(* Logix 5000 project; controller TFF vendor 1 type 14 code 107 rev 34.11; software revision 34.03; part 31 of 36 *)
(* tags used below, declared in another part *)
   FlowPath : FlowPath[64];   // Flow Path Array
   FlowPathControl : FlowPathControl;   // Flow Path Control
   Options : Options;   // Options List
   PCV001_Control : PCV_Control;   // PCV001 Control UDT
   PipeAnimation : PipeAnimation;   // HMI Pipe Animation Array
   XV001 : ALIAS FOR Valve[0];   // XV001
   XV002 : ALIAS FOR Valve[1];   // XV002
   XV003 : ALIAS FOR Valve[2];   // XV003
   XV004 : ALIAS FOR Valve[3];   // XV004
   XV005 : ALIAS FOR Valve[4];   // XV005
   XV006 : ALIAS FOR Valve[19];
   XV007 : ALIAS FOR Valve[20];
   XV401 : ALIAS FOR Valve[6];   // XV401
   XV402 : ALIAS FOR Valve[7];   // XV402
   XV403 : ALIAS FOR Valve[15];
   XV404 : ALIAS FOR Valve[16];
   XV405 : ALIAS FOR Valve[17];
   XV406 : ALIAS FOR Valve[18];
   XV411 : ALIAS FOR Valve[8];   // XV411
   XV421 : ALIAS FOR Valve[9];   // XV421
   XV431 : ALIAS FOR Valve[10];   // XV431
   XV441 : ALIAS FOR Valve[11];   // XV441
   XV901 : ALIAS FOR Valve[14];   // XV901
(* Process, continued *)

ROUTINE PipeAnimationControl   (* ladder *)
// Pipework Animation Routine
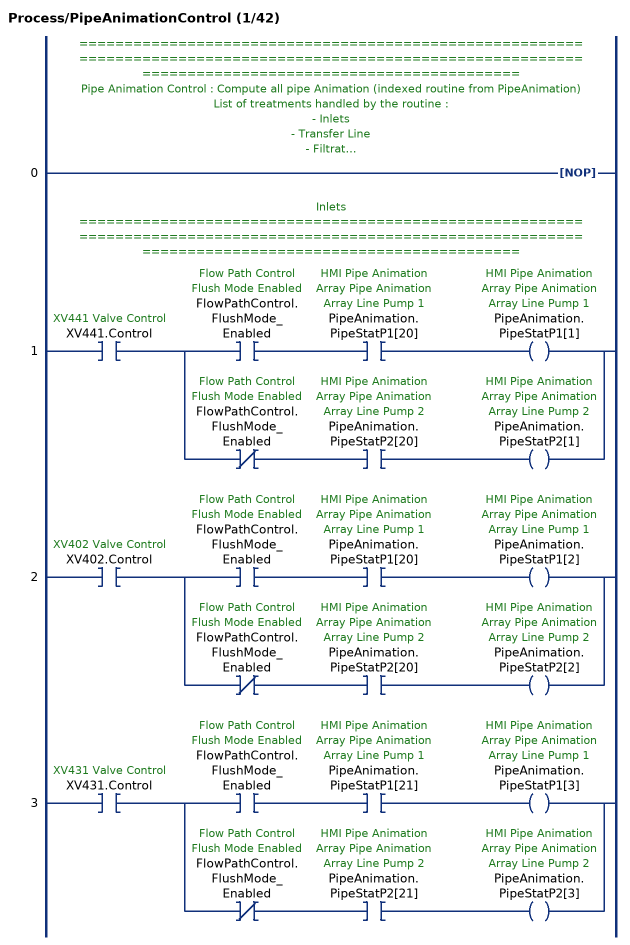
   // ==========================================================================================================================================================
   //                                                                                        Pipe Animation Control : Compute all pipe Animation (indexed routine from PipeAnimation)
   //                                                     List of treatments handled by the routine :
   //                                                          - Inlets
   //                                                          - Transfer Line
   //                                                          - Filtrate
   //                                                          - Flush
   //                                                     -----------------------------------------------------------------------------------------------------------------------------------------------------
   //                                                     History
   //                                                          2019-AUG-13 - Actemium - B. Roch - Initial version for Candidate Release 3.00.00.00.a
   //                                                          2020-OCT-01 - Merck - Q. Spindler - Modifications for Candidate Release 3.00.00.01.a
   //                                                   - Change pipe animation to add Closed Flowpath option
   // - Lock Frontal filtration flowpath
   // ========================================================================================================================================================
   0: NOP();
   // Inlets
   // ==========================================================================================================================================================
   1: XIC(XV441.Control)[XIC(FlowPathControl.FlushMode_Enabled) XIC(PipeAnimation.PipeStatP1[20]) OTE(PipeAnimation.PipeStatP1[1]) ,XIO(FlowPathControl.FlushMode_Enabled) XIC(PipeAnimation.PipeStatP2[20]) OTE(PipeAnimation.PipeStatP2[1]) ];
   2: XIC(XV402.Control)[XIC(FlowPathControl.FlushMode_Enabled) XIC(PipeAnimation.PipeStatP1[20]) OTE(PipeAnimation.PipeStatP1[2]) ,XIO(FlowPathControl.FlushMode_Enabled) XIC(PipeAnimation.PipeStatP2[20]) OTE(PipeAnimation.PipeStatP2[2]) ];
   3: XIC(XV431.Control)[XIC(FlowPathControl.FlushMode_Enabled) XIC(PipeAnimation.PipeStatP1[21]) OTE(PipeAnimation.PipeStatP1[3]) ,XIO(FlowPathControl.FlushMode_Enabled) XIC(PipeAnimation.PipeStatP2[21]) OTE(PipeAnimation.PipeStatP2[3]) ];
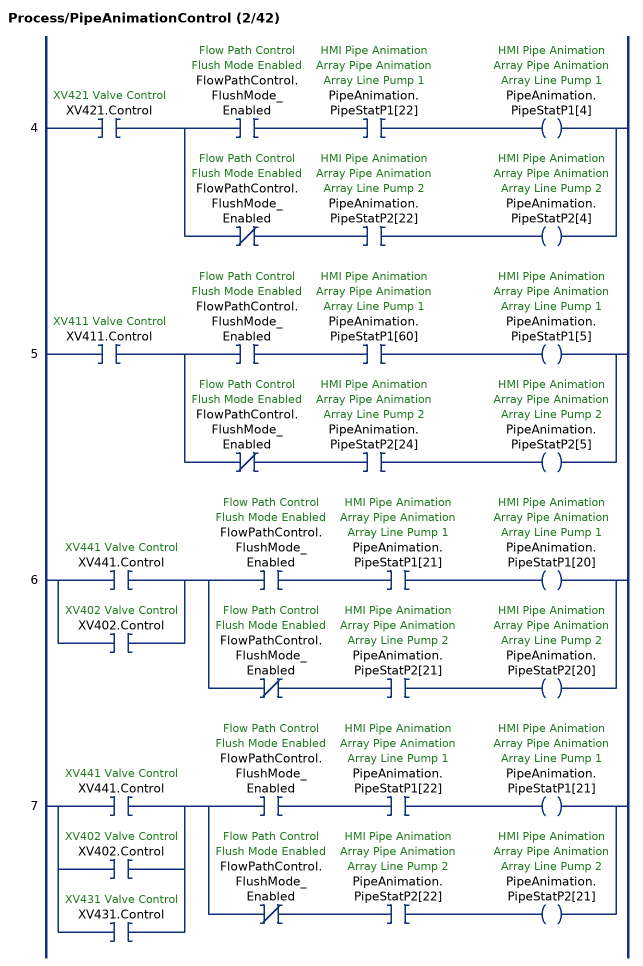
   4: XIC(XV421.Control)[XIC(FlowPathControl.FlushMode_Enabled) XIC(PipeAnimation.PipeStatP1[22]) OTE(PipeAnimation.PipeStatP1[4]) ,XIO(FlowPathControl.FlushMode_Enabled) XIC(PipeAnimation.PipeStatP2[22]) OTE(PipeAnimation.PipeStatP2[4]) ];
   5: XIC(XV411.Control)[XIC(FlowPathControl.FlushMode_Enabled) XIC(PipeAnimation.PipeStatP1[60]) OTE(PipeAnimation.PipeStatP1[5]) ,XIO(FlowPathControl.FlushMode_Enabled) XIC(PipeAnimation.PipeStatP2[24]) OTE(PipeAnimation.PipeStatP2[5]) ];
   6: [XIC(XV441.Control) ,XIC(XV402.Control) ][XIC(FlowPathControl.FlushMode_Enabled) XIC(PipeAnimation.PipeStatP1[21]) OTE(PipeAnimation.PipeStatP1[20]) ,XIO(FlowPathControl.FlushMode_Enabled) XIC(PipeAnimation.PipeStatP2[21]) OTE(PipeAnimation.PipeStatP2[20]) ];
   7: [XIC(XV441.Control) ,XIC(XV402.Control) ,XIC(XV431.Control) ][XIC(FlowPathControl.FlushMode_Enabled) XIC(PipeAnimation.PipeStatP1[22]) OTE(PipeAnimation.PipeStatP1[21]) ,XIO(FlowPathControl.FlushMode_Enabled) XIC(PipeAnimation.PipeStatP2[22]) OTE(PipeAnimation.PipeStatP2[21]) ];
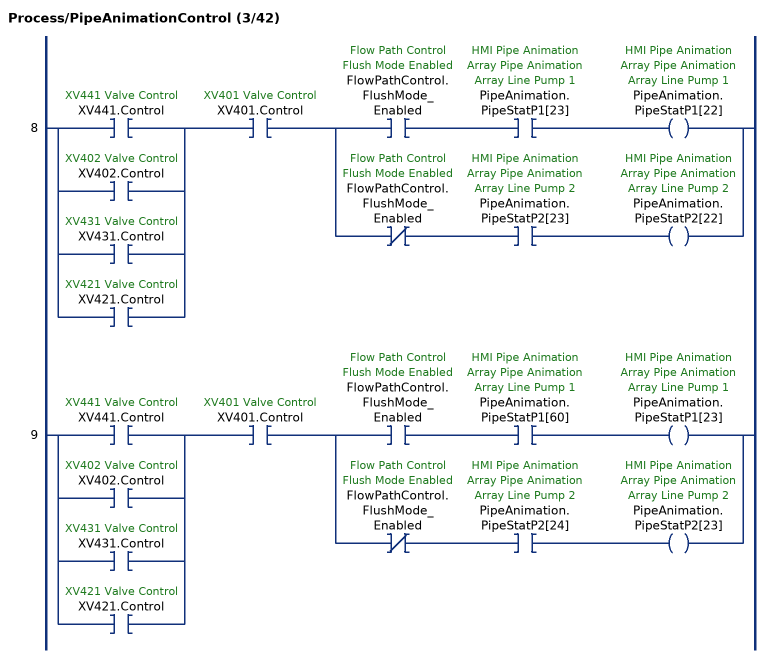
   8: [XIC(XV441.Control) ,XIC(XV402.Control) ,XIC(XV431.Control) ,XIC(XV421.Control) ]XIC(XV401.Control)[XIC(FlowPathControl.FlushMode_Enabled) XIC(PipeAnimation.PipeStatP1[23]) OTE(PipeAnimation.PipeStatP1[22]) ,XIO(FlowPathControl.FlushMode_Enabled) XIC(PipeAnimation.PipeStatP2[23]) OTE(PipeAnimation.PipeStatP2[22]) ];
   9: [XIC(XV441.Control) ,XIC(XV402.Control) ,XIC(XV431.Control) ,XIC(XV421.Control) ]XIC(XV401.Control)[XIC(FlowPathControl.FlushMode_Enabled) XIC(PipeAnimation.PipeStatP1[60]) OTE(PipeAnimation.PipeStatP1[23]) ,XIO(FlowPathControl.FlushMode_Enabled) XIC(PipeAnimation.PipeStatP2[24]) OTE(PipeAnimation.PipeStatP2[23]) ];
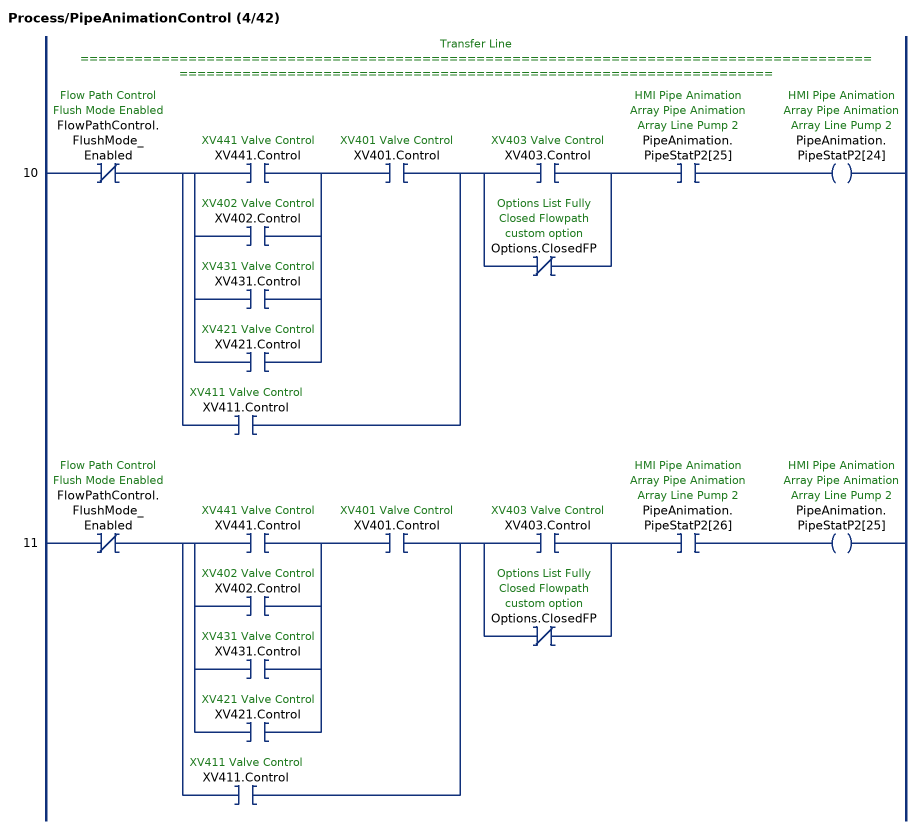
   // Transfer Line
   // ==========================================================================================================================================================
   10: XIO(FlowPathControl.FlushMode_Enabled)[[XIC(XV441.Control) ,XIC(XV402.Control) ,XIC(XV431.Control) ,XIC(XV421.Control) ] XIC(XV401.Control) ,XIC(XV411.Control) ][XIC(XV403.Control) ,XIO(Options.ClosedFP) ]XIC(PipeAnimation.PipeStatP2[25])OTE(PipeAnimation.PipeStatP2[24]);
   11: XIO(FlowPathControl.FlushMode_Enabled)[[XIC(XV441.Control) ,XIC(XV402.Control) ,XIC(XV431.Control) ,XIC(XV421.Control) ] XIC(XV401.Control) ,XIC(XV411.Control) ][XIC(XV403.Control) ,XIO(Options.ClosedFP) ]XIC(PipeAnimation.PipeStatP2[26])OTE(PipeAnimation.PipeStatP2[25]);
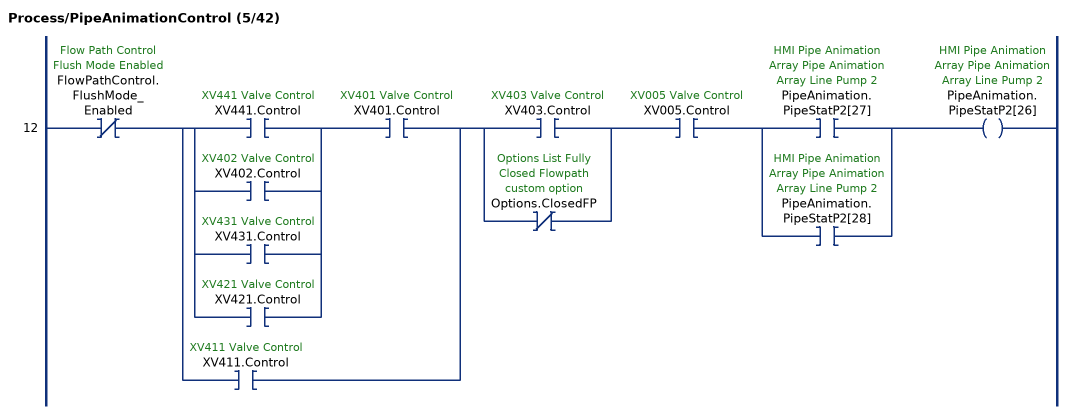
   12: XIO(FlowPathControl.FlushMode_Enabled)[[XIC(XV441.Control) ,XIC(XV402.Control) ,XIC(XV431.Control) ,XIC(XV421.Control) ] XIC(XV401.Control) ,XIC(XV411.Control) ][XIC(XV403.Control) ,XIO(Options.ClosedFP) ]XIC(XV005.Control)[XIC(PipeAnimation.PipeStatP2[27]) ,XIC(PipeAnimation.PipeStatP2[28]) ]OTE(PipeAnimation.PipeStatP2[26]);
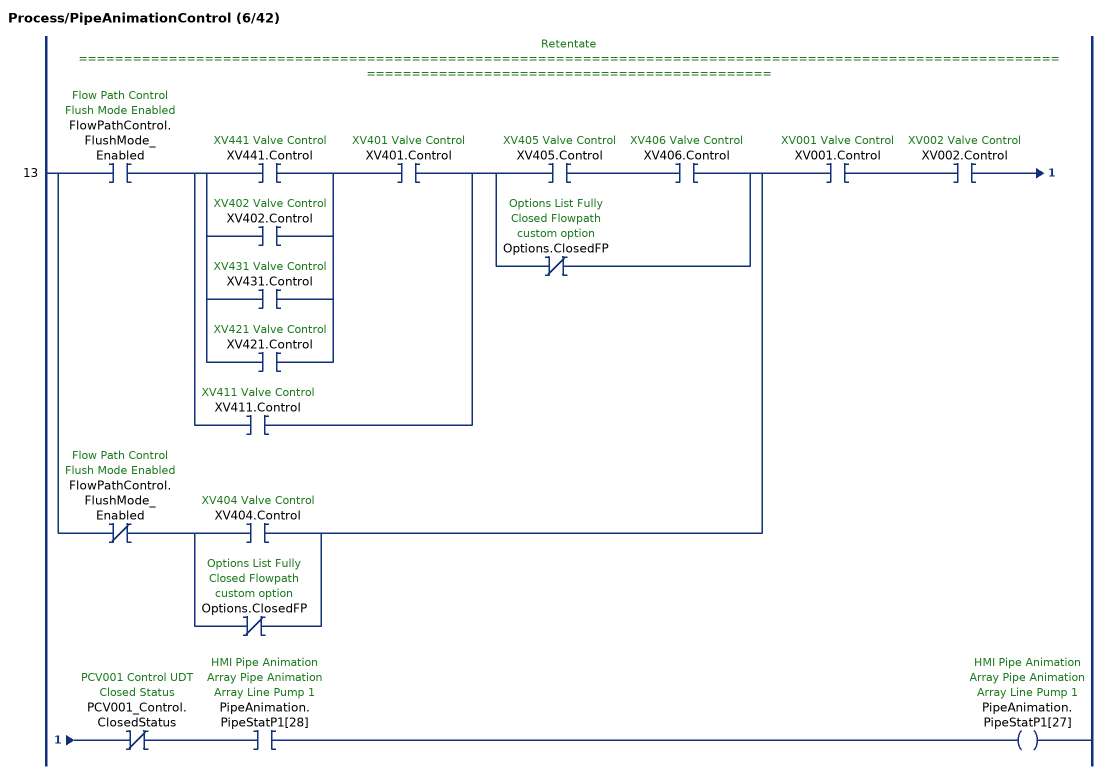
   // Retentate
   // ==========================================================================================================================================================
   13: [XIC(FlowPathControl.FlushMode_Enabled) [[XIC(XV441.Control) ,XIC(XV402.Control) ,XIC(XV431.Control) ,XIC(XV421.Control) ] XIC(XV401.Control) ,XIC(XV411.Control) ] [XIC(XV405.Control) XIC(XV406.Control) ,XIO(Options.ClosedFP) ] ,XIO(FlowPathControl.FlushMode_Enabled) [XIC(XV404.Control) ,XIO(Options.ClosedFP) ] ]XIC(XV001.Control)XIC(XV002.Control)XIO(PCV001_Control.ClosedStatus)XIC(PipeAnimation.PipeStatP1[28])OTE(PipeAnimation.PipeStatP1[27]);
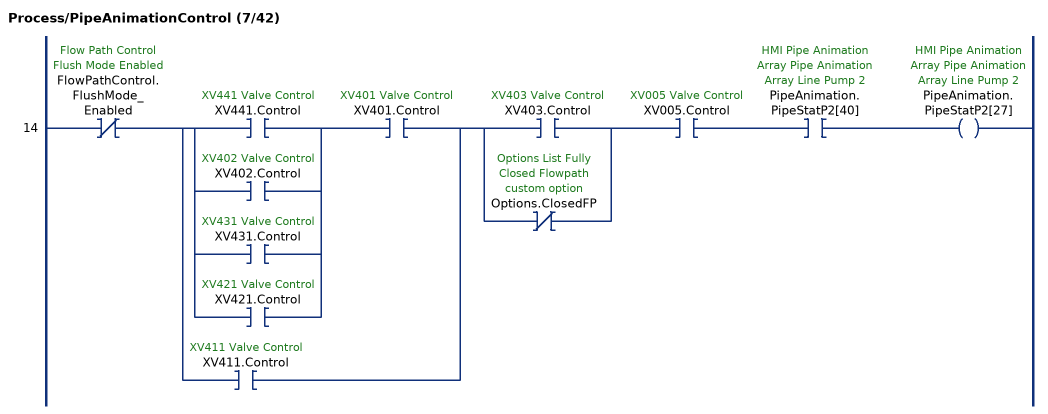
   14: XIO(FlowPathControl.FlushMode_Enabled)[[XIC(XV441.Control) ,XIC(XV402.Control) ,XIC(XV431.Control) ,XIC(XV421.Control) ] XIC(XV401.Control) ,XIC(XV411.Control) ][XIC(XV403.Control) ,XIO(Options.ClosedFP) ]XIC(XV005.Control)XIC(PipeAnimation.PipeStatP2[40])OTE(PipeAnimation.PipeStatP2[27]);
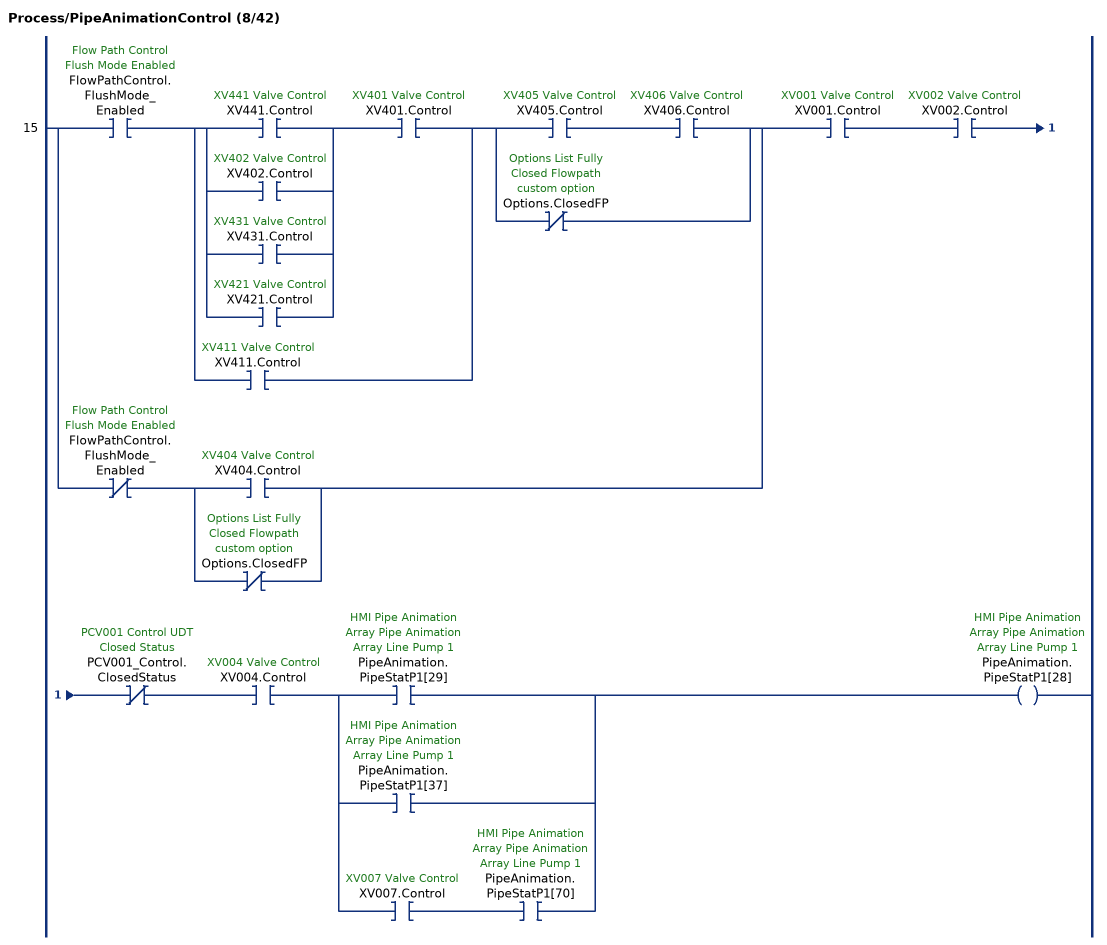
   15: [XIC(FlowPathControl.FlushMode_Enabled) [[XIC(XV441.Control) ,XIC(XV402.Control) ,XIC(XV431.Control) ,XIC(XV421.Control) ] XIC(XV401.Control) ,XIC(XV411.Control) ] [XIC(XV405.Control) XIC(XV406.Control) ,XIO(Options.ClosedFP) ] ,XIO(FlowPathControl.FlushMode_Enabled) [XIC(XV404.Control) ,XIO(Options.ClosedFP) ] ]XIC(XV001.Control)XIC(XV002.Control)XIO(PCV001_Control.ClosedStatus)XIC(XV004.Control)[[XIC(PipeAnimation.PipeStatP1[29]) ,XIC(PipeAnimation.PipeStatP1[37]) ] ,XIC(XV007.Control) XIC(PipeAnimation.PipeStatP1[70]) ]OTE(PipeAnimation.PipeStatP1[28]);
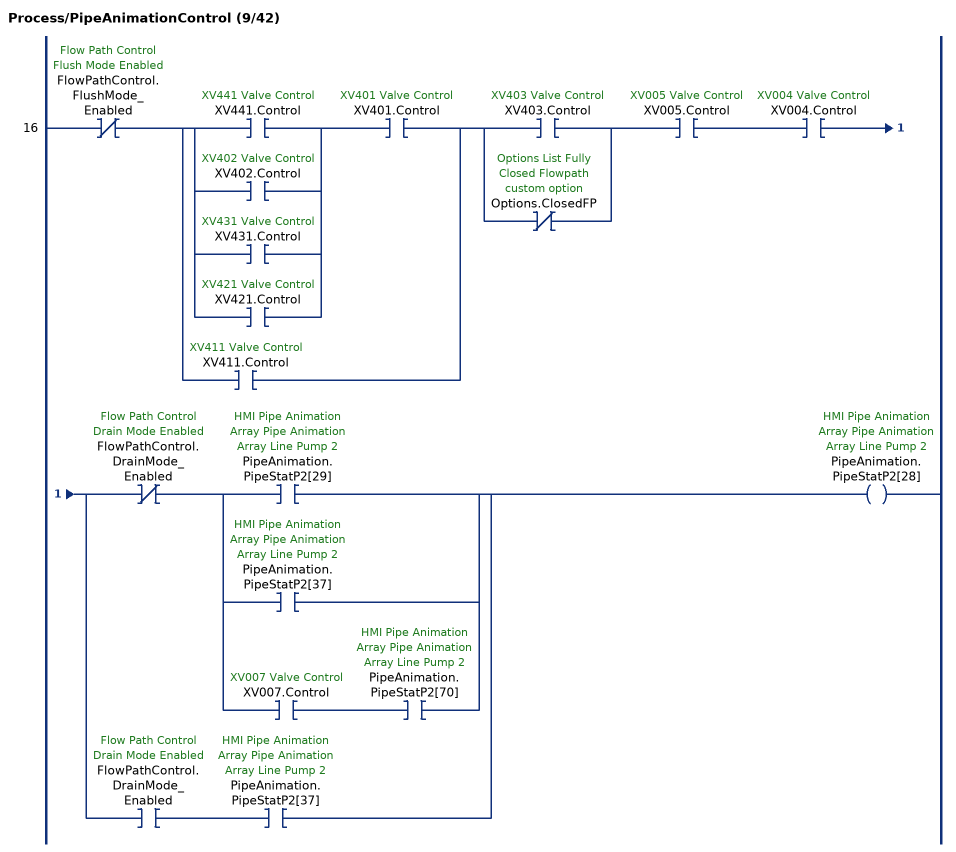
   16: XIO(FlowPathControl.FlushMode_Enabled)[[XIC(XV441.Control) ,XIC(XV402.Control) ,XIC(XV431.Control) ,XIC(XV421.Control) ] XIC(XV401.Control) ,XIC(XV411.Control) ][XIC(XV403.Control) ,XIO(Options.ClosedFP) ]XIC(XV005.Control)XIC(XV004.Control)[XIO(FlowPathControl.DrainMode_Enabled) [[XIC(PipeAnimation.PipeStatP2[29]) ,XIC(PipeAnimation.PipeStatP2[37]) ] ,XIC(XV007.Control) XIC(PipeAnimation.PipeStatP2[70]) ] ,XIC(FlowPathControl.DrainMode_Enabled) XIC(PipeAnimation.PipeStatP2[37]) ]OTE(PipeAnimation.PipeStatP2[28]);
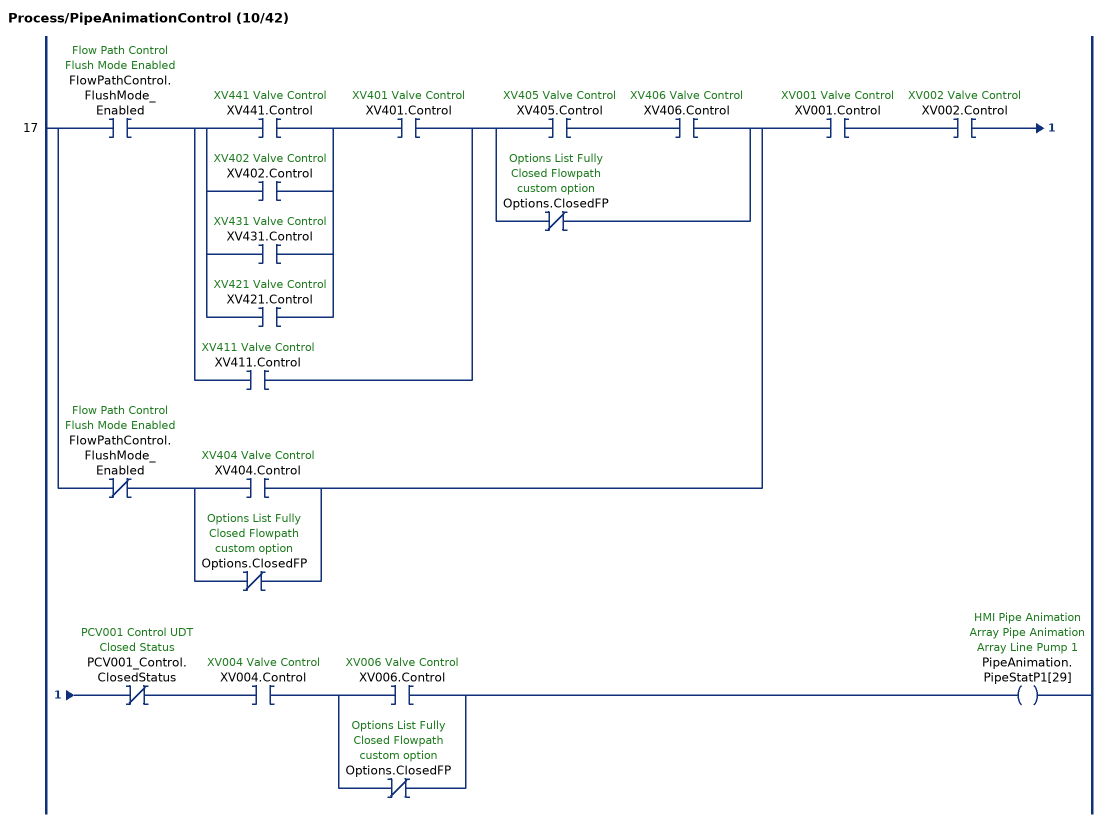
   17: [XIC(FlowPathControl.FlushMode_Enabled) [[XIC(XV441.Control) ,XIC(XV402.Control) ,XIC(XV431.Control) ,XIC(XV421.Control) ] XIC(XV401.Control) ,XIC(XV411.Control) ] [XIC(XV405.Control) XIC(XV406.Control) ,XIO(Options.ClosedFP) ] ,XIO(FlowPathControl.FlushMode_Enabled) [XIC(XV404.Control) ,XIO(Options.ClosedFP) ] ]XIC(XV001.Control)XIC(XV002.Control)XIO(PCV001_Control.ClosedStatus)XIC(XV004.Control)[XIC(XV006.Control) ,XIO(Options.ClosedFP) ]OTE(PipeAnimation.PipeStatP1[29]);
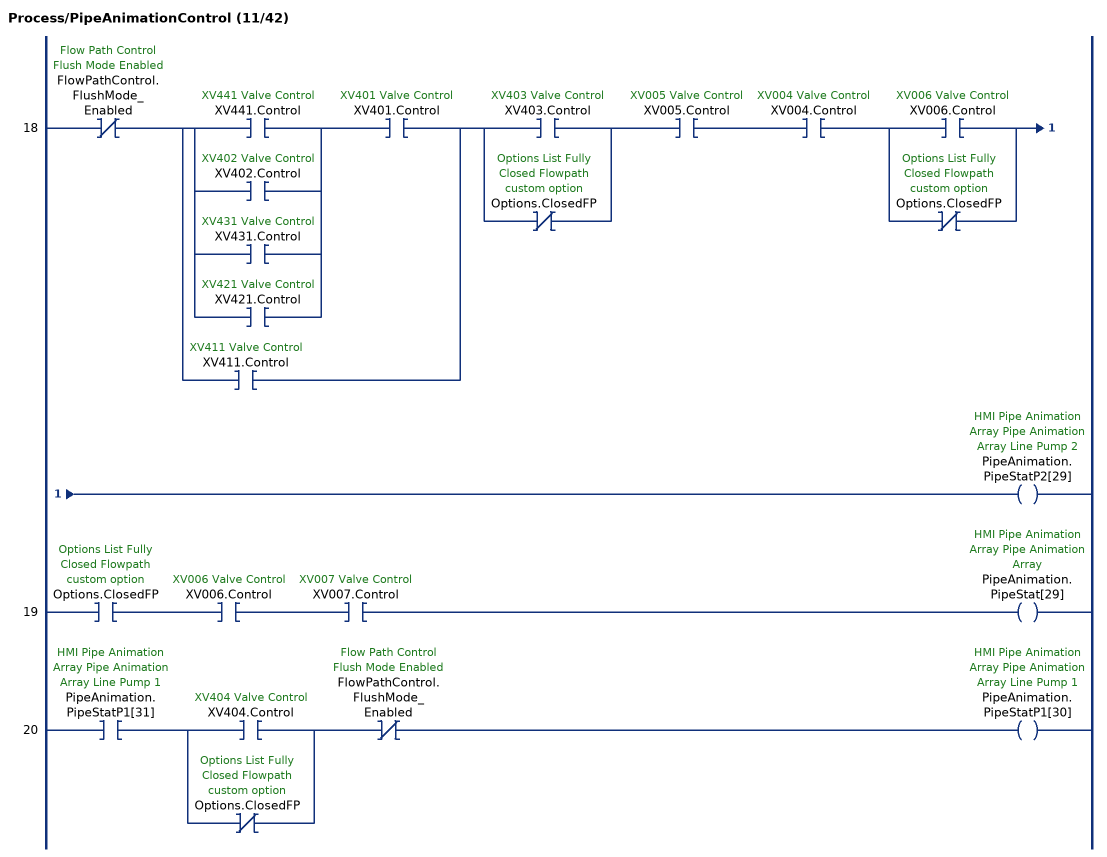
   18: XIO(FlowPathControl.FlushMode_Enabled)[[XIC(XV441.Control) ,XIC(XV402.Control) ,XIC(XV431.Control) ,XIC(XV421.Control) ] XIC(XV401.Control) ,XIC(XV411.Control) ][XIC(XV403.Control) ,XIO(Options.ClosedFP) ]XIC(XV005.Control)XIC(XV004.Control)[XIC(XV006.Control) ,XIO(Options.ClosedFP) ]OTE(PipeAnimation.PipeStatP2[29]);
   19: XIC(Options.ClosedFP)XIC(XV006.Control)XIC(XV007.Control)OTE(PipeAnimation.PipeStat[29]);
   20: XIC(PipeAnimation.PipeStatP1[31])[XIC(XV404.Control) ,XIO(Options.ClosedFP) ]XIO(FlowPathControl.FlushMode_Enabled)OTE(PipeAnimation.PipeStatP1[30]);
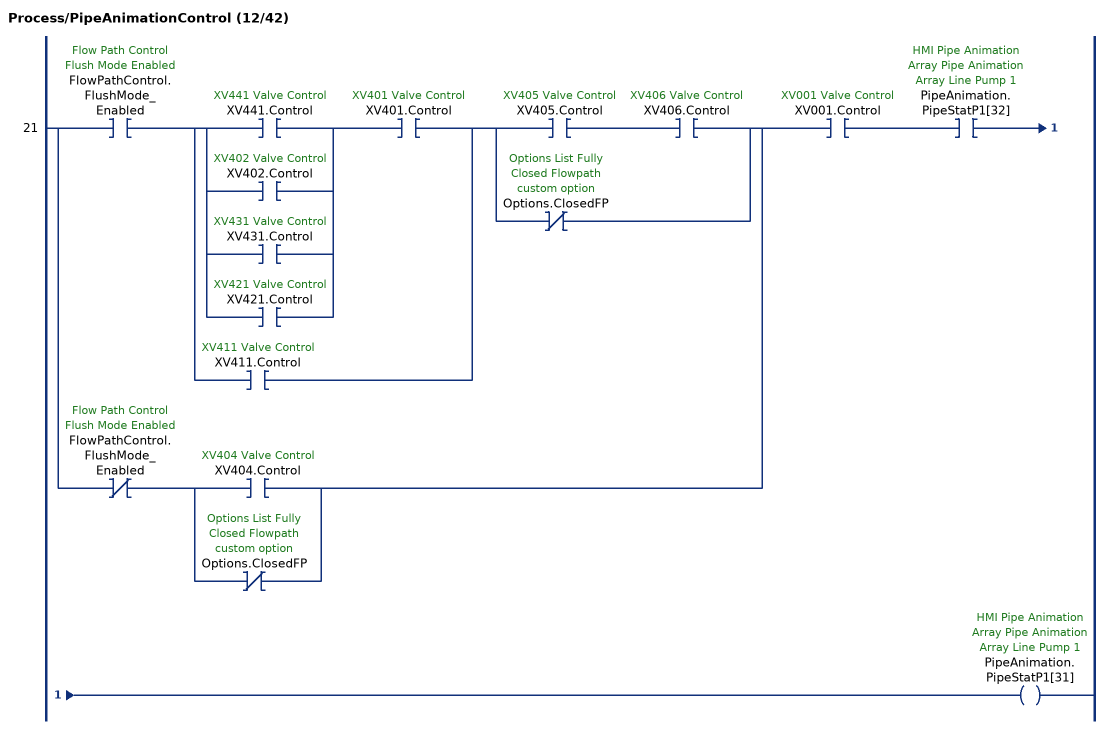
   21: [XIC(FlowPathControl.FlushMode_Enabled) [[XIC(XV441.Control) ,XIC(XV402.Control) ,XIC(XV431.Control) ,XIC(XV421.Control) ] XIC(XV401.Control) ,XIC(XV411.Control) ] [XIC(XV405.Control) XIC(XV406.Control) ,XIO(Options.ClosedFP) ] ,XIO(FlowPathControl.FlushMode_Enabled) [XIC(XV404.Control) ,XIO(Options.ClosedFP) ] ]XIC(XV001.Control)XIC(PipeAnimation.PipeStatP1[32])OTE(PipeAnimation.PipeStatP1[31]);
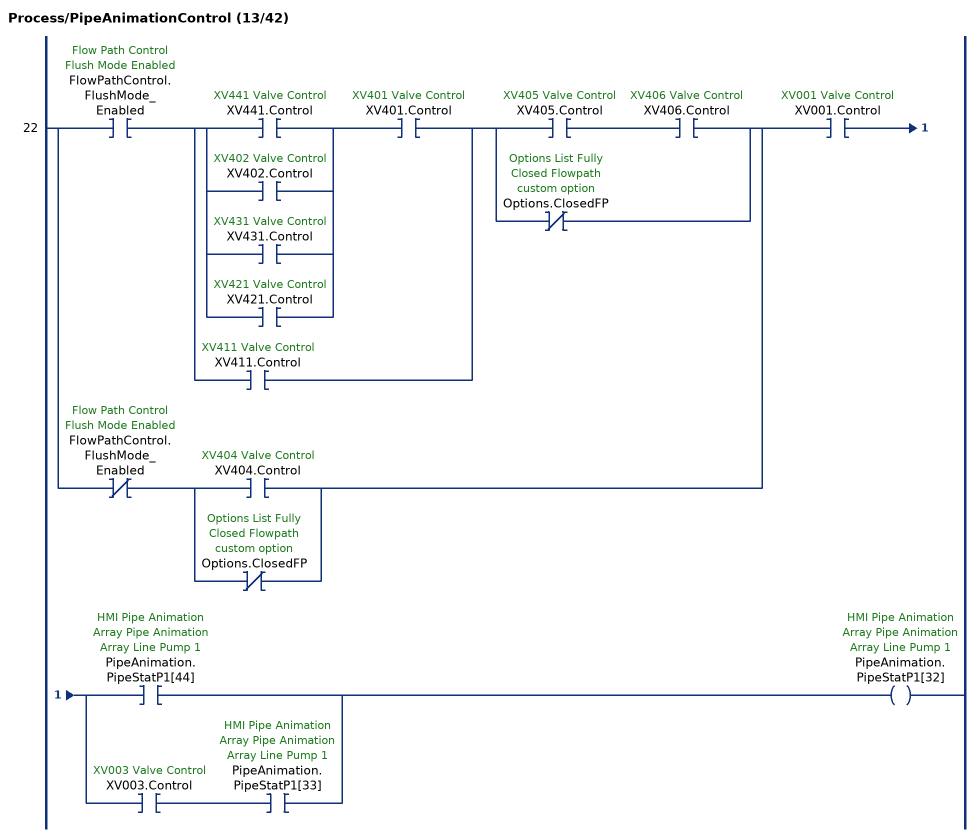
   22: [XIC(FlowPathControl.FlushMode_Enabled) [[XIC(XV441.Control) ,XIC(XV402.Control) ,XIC(XV431.Control) ,XIC(XV421.Control) ] XIC(XV401.Control) ,XIC(XV411.Control) ] [XIC(XV405.Control) XIC(XV406.Control) ,XIO(Options.ClosedFP) ] ,XIO(FlowPathControl.FlushMode_Enabled) [XIC(XV404.Control) ,XIO(Options.ClosedFP) ] ]XIC(XV001.Control)[XIC(PipeAnimation.PipeStatP1[44]) ,XIC(XV003.Control) XIC(PipeAnimation.PipeStatP1[33]) ]OTE(PipeAnimation.PipeStatP1[32]);
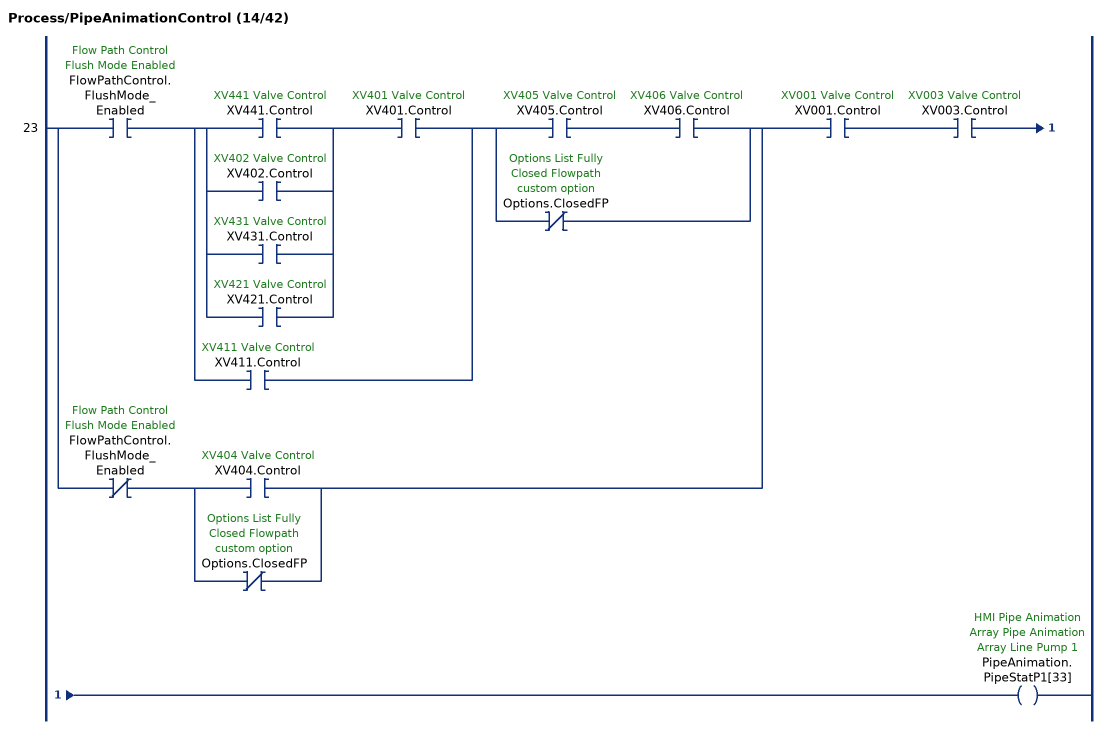
   23: [XIC(FlowPathControl.FlushMode_Enabled) [[XIC(XV441.Control) ,XIC(XV402.Control) ,XIC(XV431.Control) ,XIC(XV421.Control) ] XIC(XV401.Control) ,XIC(XV411.Control) ] [XIC(XV405.Control) XIC(XV406.Control) ,XIO(Options.ClosedFP) ] ,XIO(FlowPathControl.FlushMode_Enabled) [XIC(XV404.Control) ,XIO(Options.ClosedFP) ] ]XIC(XV001.Control)XIC(XV003.Control)OTE(PipeAnimation.PipeStatP1[33]);
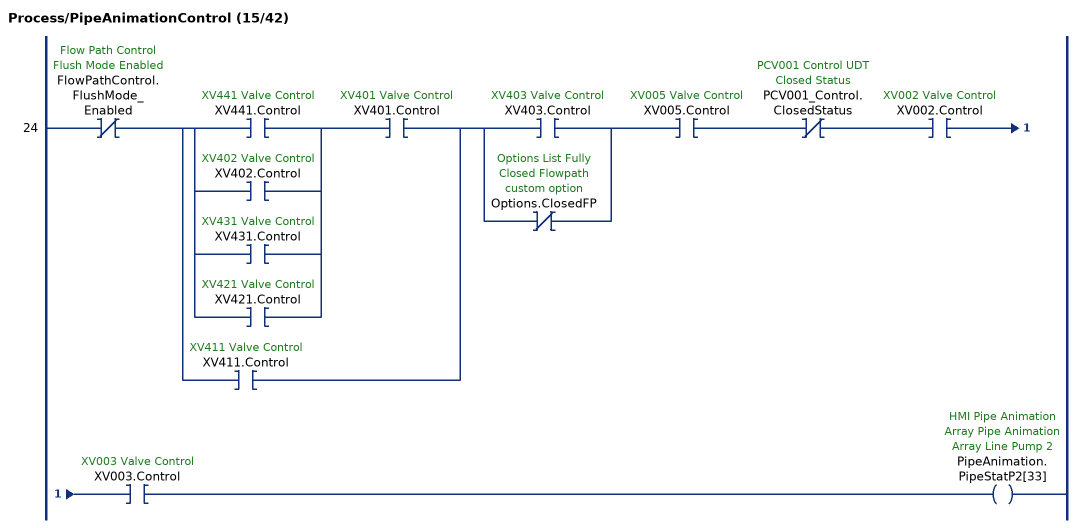
   24: XIO(FlowPathControl.FlushMode_Enabled)[[XIC(XV441.Control) ,XIC(XV402.Control) ,XIC(XV431.Control) ,XIC(XV421.Control) ] XIC(XV401.Control) ,XIC(XV411.Control) ][XIC(XV403.Control) ,XIO(Options.ClosedFP) ]XIC(XV005.Control)XIO(PCV001_Control.ClosedStatus)XIC(XV002.Control)XIC(XV003.Control)OTE(PipeAnimation.PipeStatP2[33]);
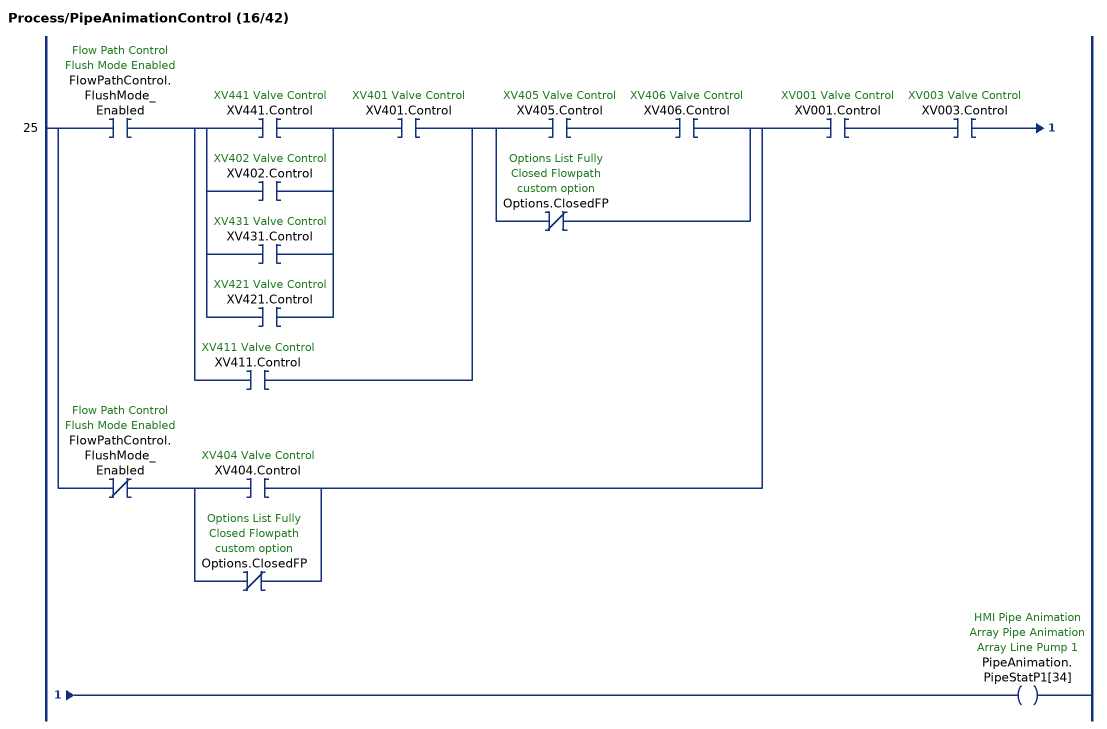
   25: [XIC(FlowPathControl.FlushMode_Enabled) [[XIC(XV441.Control) ,XIC(XV402.Control) ,XIC(XV431.Control) ,XIC(XV421.Control) ] XIC(XV401.Control) ,XIC(XV411.Control) ] [XIC(XV405.Control) XIC(XV406.Control) ,XIO(Options.ClosedFP) ] ,XIO(FlowPathControl.FlushMode_Enabled) [XIC(XV404.Control) ,XIO(Options.ClosedFP) ] ]XIC(XV001.Control)XIC(XV003.Control)OTE(PipeAnimation.PipeStatP1[34]);
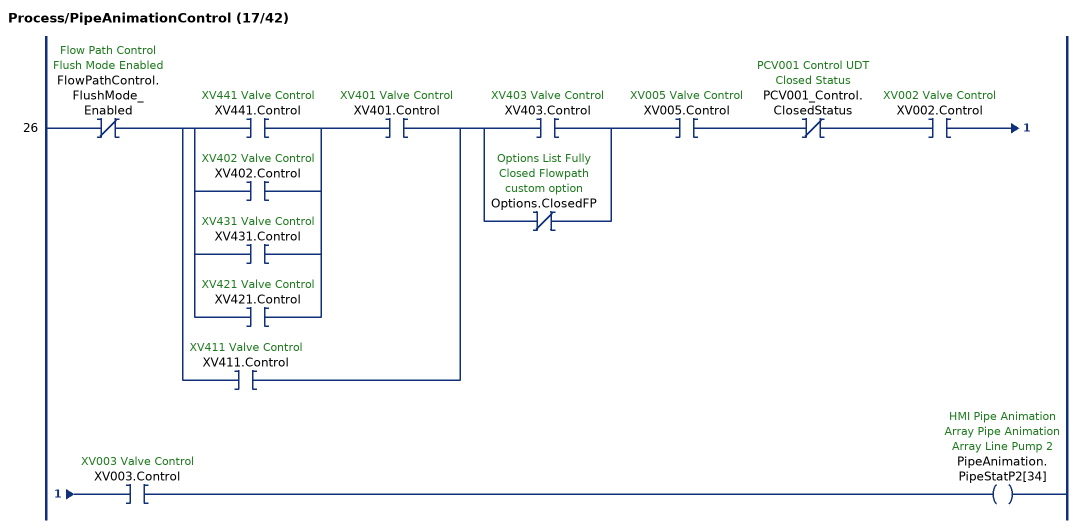
   26: XIO(FlowPathControl.FlushMode_Enabled)[[XIC(XV441.Control) ,XIC(XV402.Control) ,XIC(XV431.Control) ,XIC(XV421.Control) ] XIC(XV401.Control) ,XIC(XV411.Control) ][XIC(XV403.Control) ,XIO(Options.ClosedFP) ]XIC(XV005.Control)XIO(PCV001_Control.ClosedStatus)XIC(XV002.Control)XIC(XV003.Control)OTE(PipeAnimation.PipeStatP2[34]);
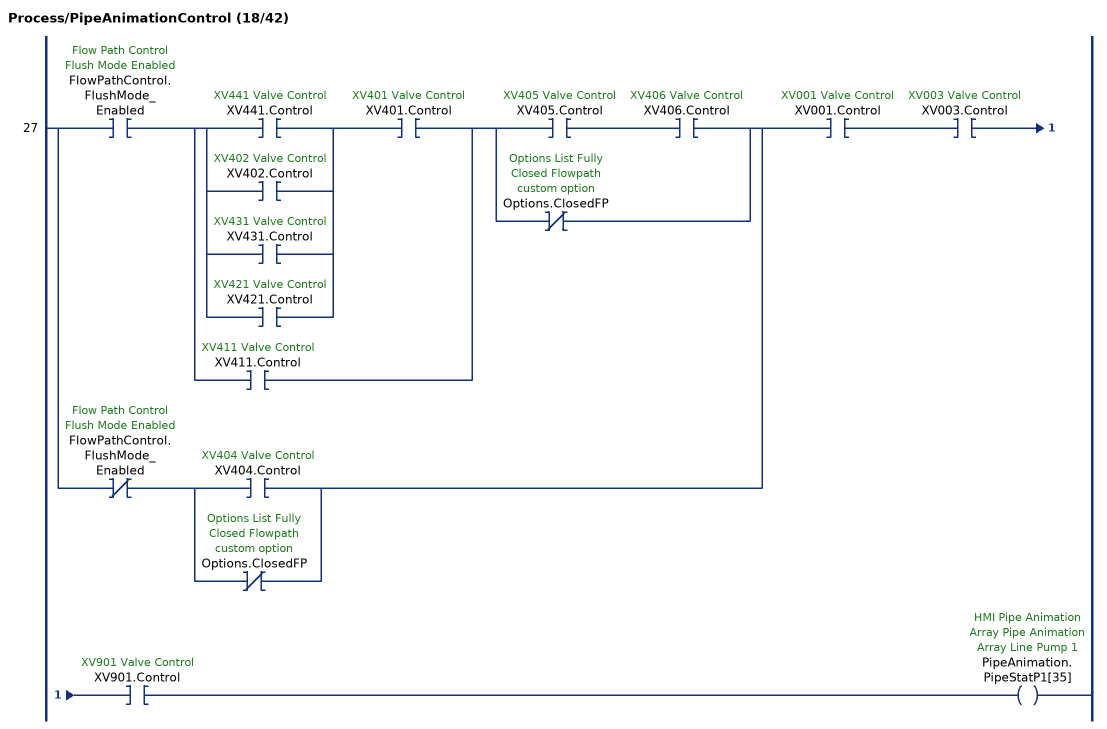
   27: [XIC(FlowPathControl.FlushMode_Enabled) [[XIC(XV441.Control) ,XIC(XV402.Control) ,XIC(XV431.Control) ,XIC(XV421.Control) ] XIC(XV401.Control) ,XIC(XV411.Control) ] [XIC(XV405.Control) XIC(XV406.Control) ,XIO(Options.ClosedFP) ] ,XIO(FlowPathControl.FlushMode_Enabled) [XIC(XV404.Control) ,XIO(Options.ClosedFP) ] ]XIC(XV001.Control)XIC(XV003.Control)XIC(XV901.Control)OTE(PipeAnimation.PipeStatP1[35]);
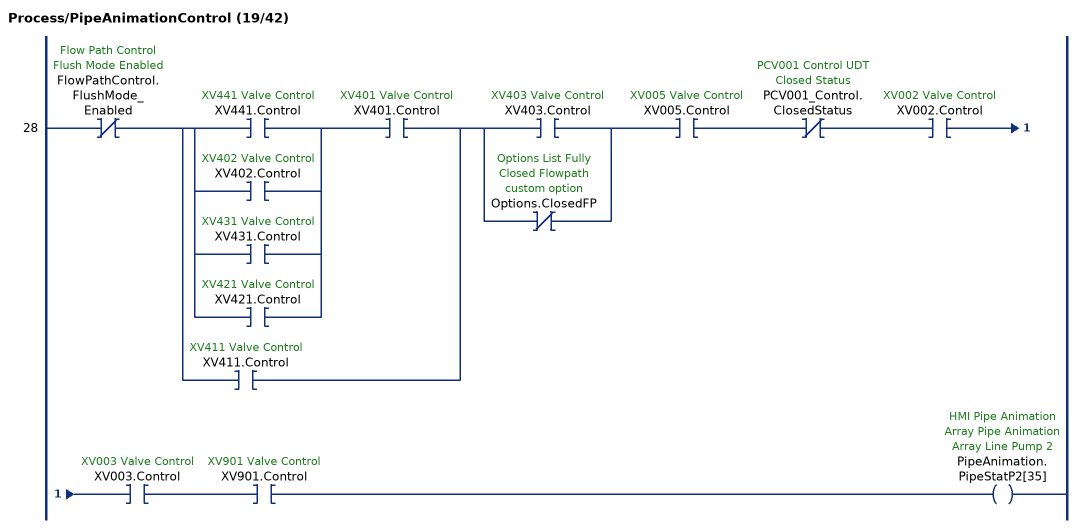
   28: XIO(FlowPathControl.FlushMode_Enabled)[[XIC(XV441.Control) ,XIC(XV402.Control) ,XIC(XV431.Control) ,XIC(XV421.Control) ] XIC(XV401.Control) ,XIC(XV411.Control) ][XIC(XV403.Control) ,XIO(Options.ClosedFP) ]XIC(XV005.Control)XIO(PCV001_Control.ClosedStatus)XIC(XV002.Control)XIC(XV003.Control)XIC(XV901.Control)OTE(PipeAnimation.PipeStatP2[35]);
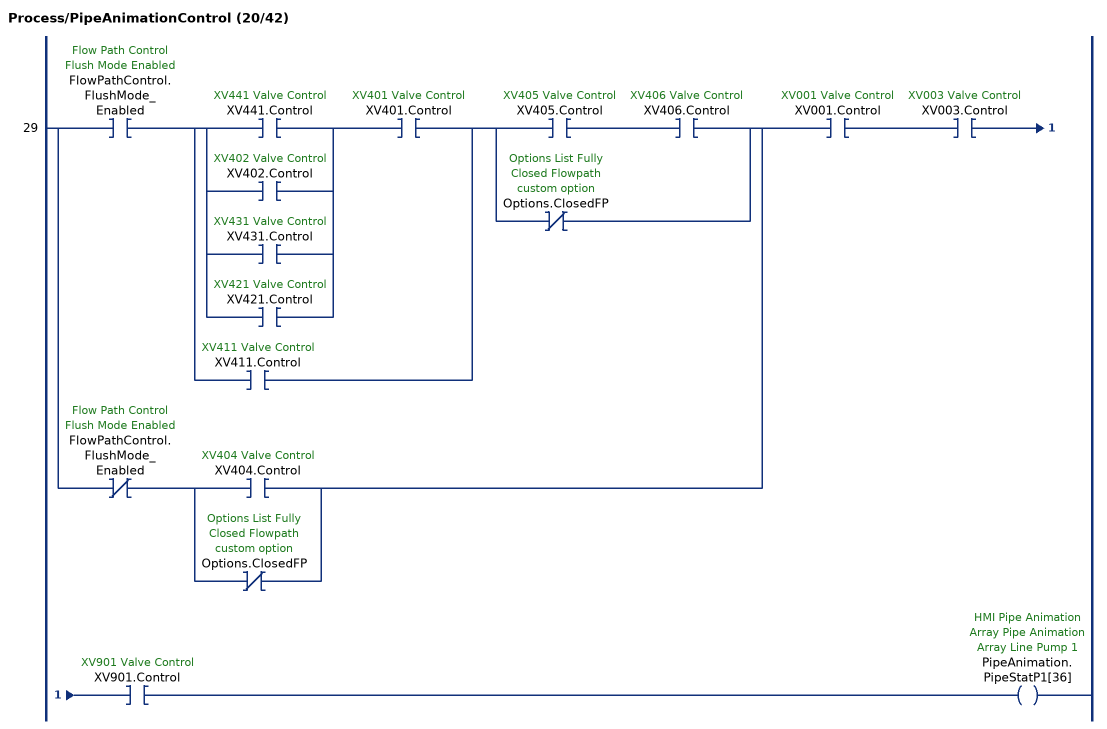
   29: [XIC(FlowPathControl.FlushMode_Enabled) [[XIC(XV441.Control) ,XIC(XV402.Control) ,XIC(XV431.Control) ,XIC(XV421.Control) ] XIC(XV401.Control) ,XIC(XV411.Control) ] [XIC(XV405.Control) XIC(XV406.Control) ,XIO(Options.ClosedFP) ] ,XIO(FlowPathControl.FlushMode_Enabled) [XIC(XV404.Control) ,XIO(Options.ClosedFP) ] ]XIC(XV001.Control)XIC(XV003.Control)XIC(XV901.Control)OTE(PipeAnimation.PipeStatP1[36]);
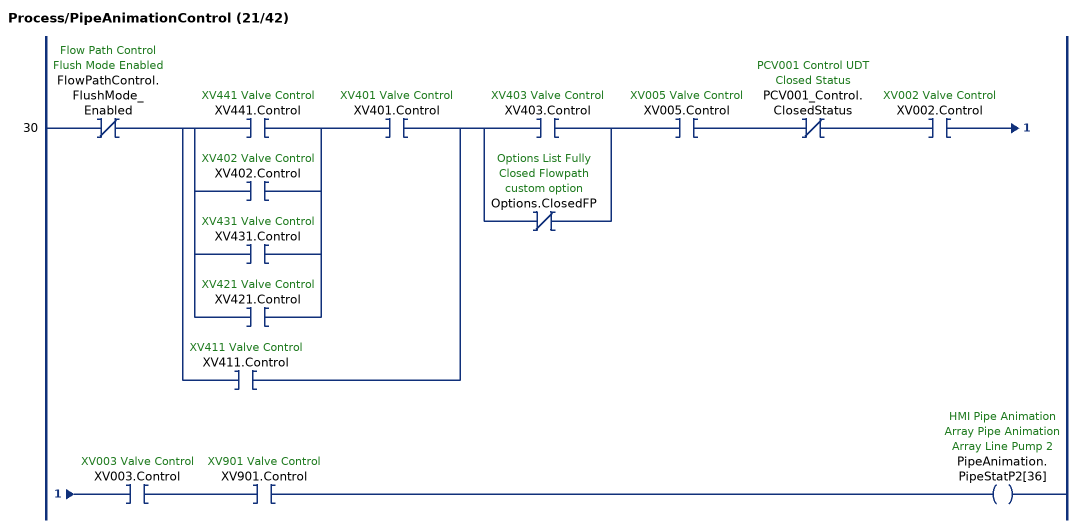
   30: XIO(FlowPathControl.FlushMode_Enabled)[[XIC(XV441.Control) ,XIC(XV402.Control) ,XIC(XV431.Control) ,XIC(XV421.Control) ] XIC(XV401.Control) ,XIC(XV411.Control) ][XIC(XV403.Control) ,XIO(Options.ClosedFP) ]XIC(XV005.Control)XIO(PCV001_Control.ClosedStatus)XIC(XV002.Control)XIC(XV003.Control)XIC(XV901.Control)OTE(PipeAnimation.PipeStatP2[36]);
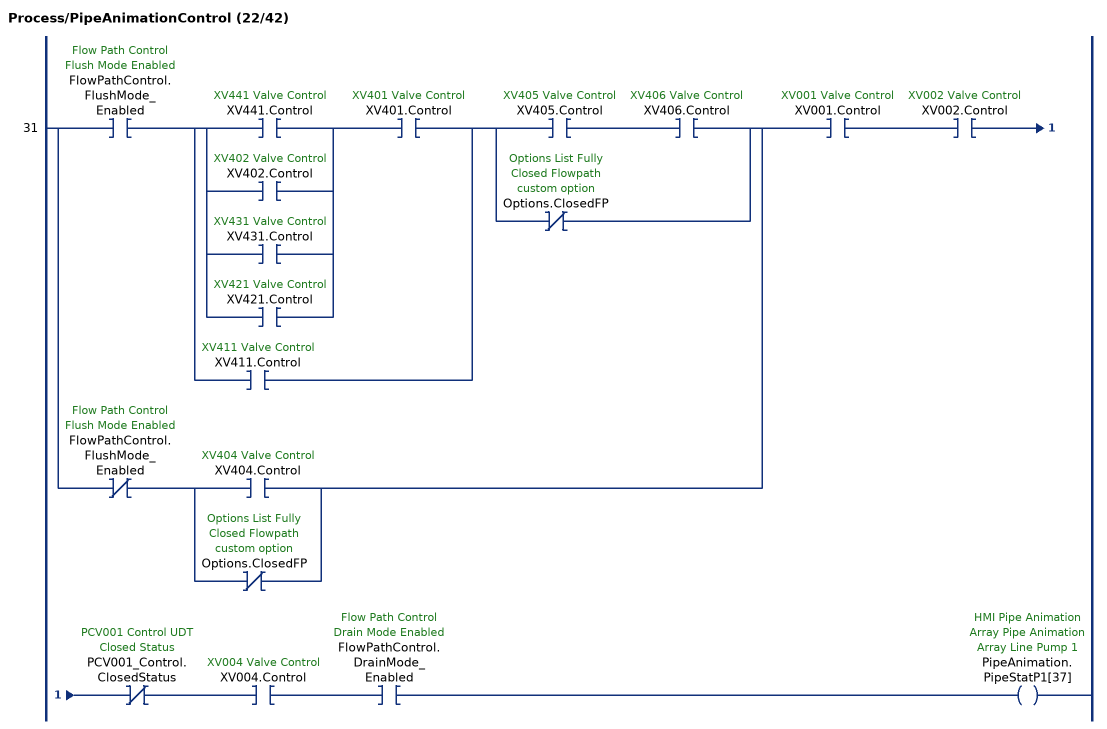
   31: [XIC(FlowPathControl.FlushMode_Enabled) [[XIC(XV441.Control) ,XIC(XV402.Control) ,XIC(XV431.Control) ,XIC(XV421.Control) ] XIC(XV401.Control) ,XIC(XV411.Control) ] [XIC(XV405.Control) XIC(XV406.Control) ,XIO(Options.ClosedFP) ] ,XIO(FlowPathControl.FlushMode_Enabled) [XIC(XV404.Control) ,XIO(Options.ClosedFP) ] ]XIC(XV001.Control)XIC(XV002.Control)XIO(PCV001_Control.ClosedStatus)XIC(XV004.Control)XIC(FlowPathControl.DrainMode_Enabled)OTE(PipeAnimation.PipeStatP1[37]);
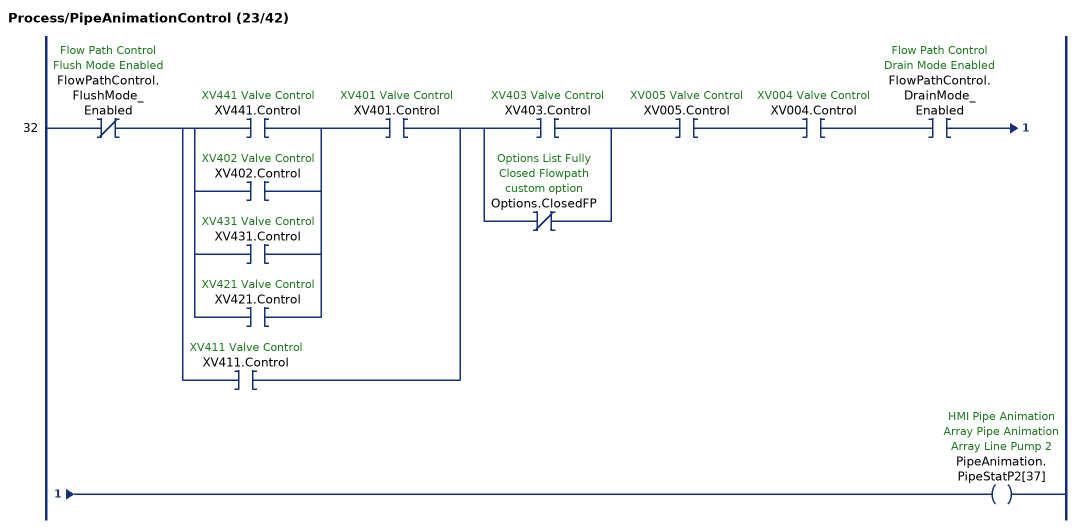
   32: XIO(FlowPathControl.FlushMode_Enabled)[[XIC(XV441.Control) ,XIC(XV402.Control) ,XIC(XV431.Control) ,XIC(XV421.Control) ] XIC(XV401.Control) ,XIC(XV411.Control) ][XIC(XV403.Control) ,XIO(Options.ClosedFP) ]XIC(XV005.Control)XIC(XV004.Control)XIC(FlowPathControl.DrainMode_Enabled)OTE(PipeAnimation.PipeStatP2[37]);
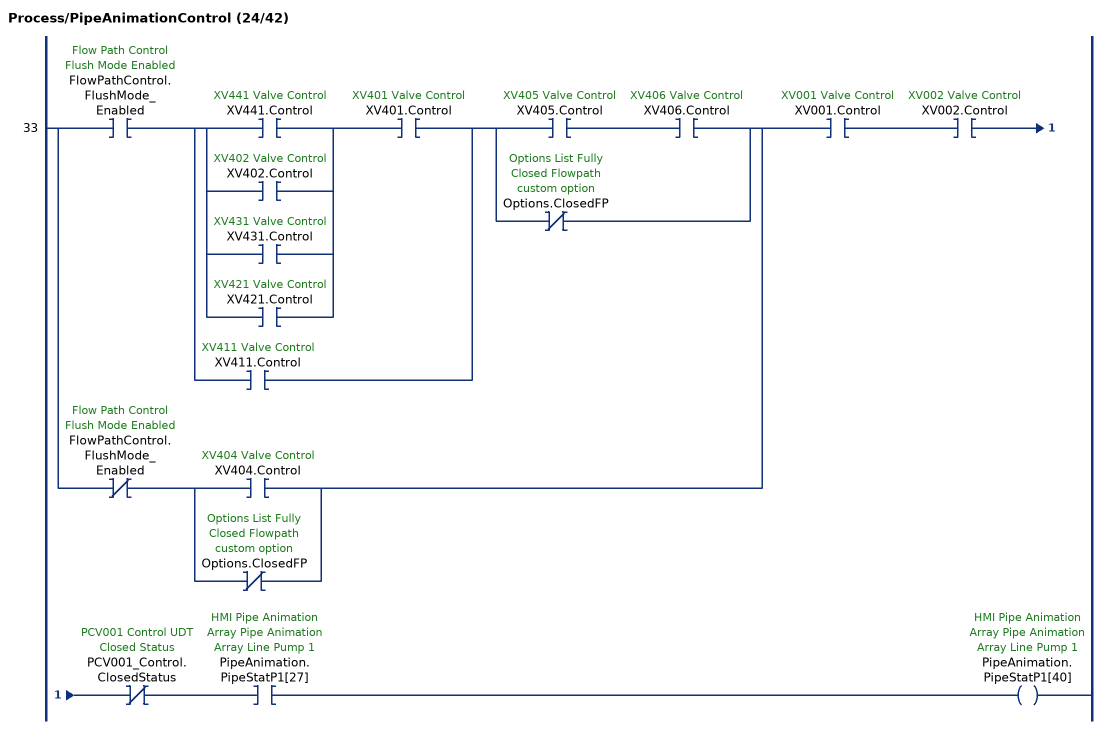
   33: [XIC(FlowPathControl.FlushMode_Enabled) [[XIC(XV441.Control) ,XIC(XV402.Control) ,XIC(XV431.Control) ,XIC(XV421.Control) ] XIC(XV401.Control) ,XIC(XV411.Control) ] [XIC(XV405.Control) XIC(XV406.Control) ,XIO(Options.ClosedFP) ] ,XIO(FlowPathControl.FlushMode_Enabled) [XIC(XV404.Control) ,XIO(Options.ClosedFP) ] ]XIC(XV001.Control)XIC(XV002.Control)XIO(PCV001_Control.ClosedStatus)XIC(PipeAnimation.PipeStatP1[27])OTE(PipeAnimation.PipeStatP1[40]);
